(* IEC 61131-3 sources: axsharp/src/ix.compiler/tests/integration/actual/lib1/src, 1 file *)

(* ---- library.st ---- *)
NAMESPACE lib1

    CLASS PUBLIC MyClass
        VAR PUBLIC
            MyString : STRING;
            MyInt : INT;
        END_VAR

        VAR PRIVATE

        END_VAR

        METHOD PUBLIC MyMethod : BOOL
            MyMethod := FALSE;
        END_METHOD
    END_CLASS

END_NAMESPACE
